// TIA Portal V21 export
// export: Created 2026-11-10T19:21:32.5304084Z, ExportSetting WithDefaults, DisplayName Totally Integrated Automation Portal, DisplayVersion V21 Update 3, DisplayName STEP 7 Professional, DisplayVersion V21 Update 3, DisplayName STEP 7 Safety, DisplayVersion V21, DisplayName Tech WebApplication, DisplayVersion V21, DisplayName WinCC Basic/Comfort/Advanced, DisplayVersion V21 Update 3, DisplayName WinCC Unified, DisplayVersion V21 Update 3
FUNCTION_BLOCK "FB_Lad_pt006"   // FB1, LAD
{ S7_Optimized_Access := 'TRUE' }
VERSION : 0.1
// stored: AutoNumber true, IsIECCheckEnabled false, IsRetainMemResEnabled false, MemoryReserve 100, SetENOAutomatically false, UDAEnableTagReadback false
   VAR_INPUT
      v_req : Bool;
      v_port : PORT;
   END_VAR
   VAR_OUTPUT
      v_done : Bool;
      v_error : Bool;
      v_status : Word;
   END_VAR
   VAR
      inst { S7_SetPoint := 'True'} : Receive_Reset;
   END_VAR
BEGIN

REGION Network 1: RCV_RST - Delete receive buffer
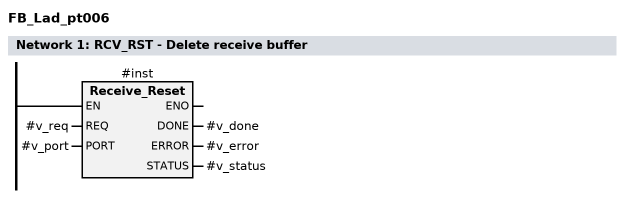
   RUNG wire#powerrail
      #inst.Receive_Reset(REQ := #v_req, PORT := #v_port, DONE => #v_done, ERROR => #v_error, STATUS => #v_status)
   END_RUNG
   // the same network as SCL:
   #inst(REQ := #v_req, PORT := #v_port, DONE => #v_done, ERROR => #v_error, STATUS => #v_status);   // Receive_Reset
END_REGION
END_FUNCTION_BLOCK
